(*
SPDX-FileCopyrightText: © 2026 Oleksandr Tiutyk <trofimich@gmail.com>
SPDX-License-Identifier: MIT
License: https://opensource.org/license/mit
*)

(*!
<summary>
Beckhoff bidirectional incremental encoder channel process image.
</summary>
<description>
Aggregates input position/status/latch and output control/preset for an incremental encoder interface.
Requires the matching 32-bit EL5101 enhanced or EL5151 main PDOs. EL5152 uses the latch-free
INCREMENTAL_ENCODER_COUNTER_CHANNEL; do not substitute these channel types for each other.
When used for I/O, link located fields or their containing buffers to the matching selected PDOs.
The record is not a packed wire buffer; compiler padding is not part of the device specification.
Unlinked/default values do not prove valid I/O. The caller evaluates bus/channel validity before use.
Use one owner task per instance and externally synchronize other access; multi-field snapshots are not atomic.
Copies store data without creating hardware links. Keep borrowed field references valid while consumers are bound.
This passive record performs no validation, synchronization, configuration or protocol advancement.
</description>
*)
TYPE INCREMENTAL_ENCODER_CHANNEL :
STRUCT
	In : INCREMENTAL_ENCODER_INPUT_CHANNEL;
	Out : INCREMENTAL_ENCODER_OUTPUT_CHANNEL;
END_STRUCT
END_TYPE

(* stored: Version 1.1.0.1, ProductVersion 3.1.4026.20
   DUT INCREMENTAL_ENCODER_CHANNEL: Id {e60b5e74-037a-4705-84f0-571ee29612ac} *)
